(* CODESYS project Tc3_McCoordinatedMotion.library
   TcLibraryId: Beckhoff Automation GmbH|Tc3_McCoordinatedMotion|4.0.17.0
   Company: Beckhoff Automation GmbH
   Title: Tc3_McCoordinatedMotion
   Placeholder: Tc3_McCoordinatedMotion
   Version: 4.0.17.0

Project tree, tasks and I/O mapping:
  libraries: Tc2_MC2, * (Beckhoff Automation GmbH); Tc3_Mc3Definitions, 4.0.17.0 (Beckhoff Automation GmbH); Tc3_Physics, 4.0.17.0 (Beckhoff Automation GmbH)
  POUs/
    Administrative/
      function ACSIDX_TO_IDENTINGROUP [ST]
      function MCSAXISTYPE_TO_IDENTINGROUP [ST]
      function MCSIDX_TO_IDENTINGROUP [ST]
      function block MC_AddAxisToGroup [ST]: FB_init, FB_exit
      function block MC_GroupDisable [ST]: FB_init, FB_exit
      function block MC_GroupEnable [ST]: FB_init, FB_exit
      function block MC_GroupReadError [ST]: FB_init, FB_exit
      function block MC_GroupReadStatus [ST]: FB_init, FB_exit
      function block MC_GroupReadTrajectoryInformation [ST]: FB_init, FB_exit
      function block MC_GroupReset [ST]: FB_init, FB_exit
      function block MC_GroupSetOverride [ST]: FB_init, FB_exit
      function block MC_GroupSetSetpointSource [ST]: FB_init, FB_exit
      function block MC_RemoveAxisFromGroup [ST]: FB_init, FB_exit
      function block MC_SetCoordinateTransform [ST]: FB_init, FB_exit
      function block MC_SetCoordinateTransformPreparation [ST]: FB_init, FB_exit
      function block MC_TrackConveyorBelt [ST]: FB_init, FB_exit
      function block MC_UngroupAllAxes [ST]: FB_init, FB_exit
      function UDINT_TO_IDENTINGROUP [ST]
    Motion/
      function block MC_MovePath [ST]: FB_init, FB_exit
      function block MC_BlockerPreparation [ST]: FB_init, FB_exit
      function block MC_DwellTimePreparation [ST]: FB_init, FB_exit
      function block MC_GroupHalt [ST]: FB_init, FB_exit
      function block MC_GroupStop [ST]: FB_init, FB_exit
      function block MC_MoveBlendingPreparation [ST]: FB_init, FB_exit
      function block MC_MoveCircularAbsolutePreparation [ST]: FB_init, FB_exit
      function block MC_GroupReadBlockerStatus [ST]: FB_init, FB_exit
      function block MC_MoveDirectPreparation [ST]: FB_init, FB_exit
      function block MC_MoveLinearAbsolutePreparation [ST]: FB_init, FB_exit
      function block MC_ReleaseBlocker [ST]: FB_init, FB_exit
      function block MC_CalcTrafo [ST]: FB_init, FB_exit
  DUTs/
    function block MC_PATH_DATA_REF [ST]: ClearPath, FB_init, FB_exit
    data type AXES_GROUP_REF
    data type IDENT_IN_GROUP_REF
    Enums/
      data type MC_MCS_AXIS_TYPE
      data type MC_CIRC_MODE
      data type MC_CIRC_PATHCHOICE
      data type MC_TRANSITION_MODE
      data type ECmSetpointSource
      data type ETrackingSyncPosStrategy
    data type MC_COORD_REF
    data type MC_TRAJECTORY_ENTRY
    CalcTrafo/
      data type E_CalcTrafoMetaInfoScara
      data type E_CalcTrafoMetaInfo5DType1
      data type U_CalcTrafoMetaInfo
  GVLs/
    global variables GVL
  Version/
    global variables Global_Version
*)

// DUTs/AXES_GROUP_REF
(* Contains the information passed between Nc and Plc for each group. *)
{attribute 'TcIecLibraryType'}
{attribute 'Namespace' := 'Tc3_McCoordinatedMotion'}
TYPE AXES_GROUP_REF : 
	STRUCT
		(* Data from PLC to MC. *)
		{attribute 'GUID' := '0E2E3852-A98C-4AF3-81E2-209EE128940C'}
		{attribute 'Namespace' := 'MC'}
		PlcToNc AT %Q* : MC.CDT_PLCTOMC_GROUP;
		(* Data from MC to PLC. *)
		{attribute 'GUID' := '467F4325-10DF-4BC1-88DD-E8240EB4F8E3'}
		{attribute 'Namespace' := 'MC'}
		NcToPlc AT %I* : MC.CDT_MCTOPLC_GROUP;
	END_STRUCT
END_TYPE

// DUTs/IDENT_IN_GROUP_REF
{attribute 'TcIecLibraryType'}
{attribute 'Namespace' := 'Tc3_McCoordinatedMotion'}
TYPE IDENT_IN_GROUP_REF : Tc3_Physics.CoordinateType;
END_TYPE

// DUTs/MC_COORD_REF
{attribute 'TcIecLibraryType'}
{attribute 'Namespace' := 'Tc3_McCoordinatedMotion'}
TYPE MC_COORD_REF : GLOBAL.OTCID;
END_TYPE

// DUTs/MC_TRAJECTORY_ENTRY
{attribute 'TcIecLibraryType'}
{attribute 'Namespace' := 'Tc3_McCoordinatedMotion'}
TYPE MC_TRAJECTORY_ENTRY : 
	STRUCT
		InvokeId : UDINT;
		Active : BOOL;
		 {attribute 'hide'}
		_reserved1 : ARRAY [1..3] OF USINT;
		RemainingCartesianLength : LREAL;
		RemainingDuration : LREAL;
	END_STRUCT
END_TYPE

// DUTs/Enums/MC_MCS_AXIS_TYPE
{attribute 'TcIecLibraryType'}
{attribute 'Namespace' := 'Tc3_McCoordinatedMotion'}
{attribute 'hide'}
TYPE MC_MCS_AXIS_TYPE : (mcAxisTypeMcsX:=17, mcAxisTypeMcsY:=33, mcAxisTypeMcsZ:=49, mcAxisTypeMcsA1:=65, mcAxisTypeMcsA2:=66, mcAxisTypeMcsA3:=67, mcAxisTypeMcsB1:=81, mcAxisTypeMcsB2:=82, mcAxisTypeMcsB3:=83, mcAxisTypeMcsC1:=97, mcAxisTypeMcsC2:=98, mcAxisTypeMcsC3:=99) UDINT;
END_TYPE

// DUTs/Enums/MC_CIRC_MODE
{attribute 'TcIecLibraryType'}
{attribute 'Namespace' := 'Tc3_McCoordinatedMotion'}
TYPE MC_CIRC_MODE : (mcCircModeInvalid:=0, mcCircModeBorder:=8192, mcCircModeCenter:=8193, mcCircModeRadius:=8194) UINT;
END_TYPE

// DUTs/Enums/MC_CIRC_PATHCHOICE
{attribute 'TcIecLibraryType'}
{attribute 'Namespace' := 'Tc3_McCoordinatedMotion'}
TYPE MC_CIRC_PATHCHOICE : (mcCircPathChoiceClockwise:=12288, mcCircPathChoiceCounterClockwise:=12289, mcCircPathChoiceShortSegment:=12290, mcCircPathChoiceLongSegment:=12291) UINT;
END_TYPE

// DUTs/Enums/MC_TRANSITION_MODE
{attribute 'TcIecLibraryType'}
{attribute 'Namespace' := 'Tc3_McCoordinatedMotion'}
TYPE MC_TRANSITION_MODE : (mcTransModeNone:=4096, mcTransModeStartVelocity:=4097, mcTransModeConstantVelocity:=4098, mcTransModeCornerDistance:=4099, mcTransModeMaxCornerDeviation:=4100, mcTransModeCornerDistanceAdvanced:=4106) UINT;
END_TYPE

// DUTs/Enums/ECmSetpointSource
{attribute 'TcIecLibraryType'}
{attribute 'Namespace' := 'Tc3_McCoordinatedMotion'}
{attribute 'qualified_only'}
TYPE ECmSetpointSource : (Group:=1, MCS:=2, ACS:=3) UINT;
END_TYPE

// DUTs/Enums/ETrackingSyncPosStrategy
{attribute 'TcIecLibraryType'}
{attribute 'Namespace' := 'Tc3_McCoordinatedMotion'}
{attribute 'hide'}
{attribute 'qualified_only'}
TYPE ETrackingSyncPosStrategy : (FastestSync:=0, ObjectPos:=1) UINT;
END_TYPE

// DUTs/CalcTrafo/E_CalcTrafoMetaInfoScara
{attribute 'TcIecLibraryType'}
{attribute 'Namespace' := 'Tc3_McCoordinatedMotion'}
TYPE E_CalcTrafoMetaInfoScara : (scaraLeftArm:=1, scaraRightArm:=2, scaraActualConfig:=3) WORD;
END_TYPE

// DUTs/CalcTrafo/E_CalcTrafoMetaInfo5DType1
{attribute 'TcIecLibraryType'}
{attribute 'Namespace' := 'Tc3_McCoordinatedMotion'}
TYPE E_CalcTrafoMetaInfo5DType1 : (
	d5Type1Quad14:=1, 	(* M3: -90..90 and TCP in same quadrants *)
	d5Type1Quad23:=2, 	(* M3: -90..90 and TCP OUTSIDE these quadrants *)
	d5Type1ActualConfig:=3
) WORD;
END_TYPE

// DUTs/CalcTrafo/U_CalcTrafoMetaInfo
{attribute 'TcIecLibraryType'}
{attribute 'Namespace' := 'Tc3_McCoordinatedMotion'}
TYPE U_CalcTrafoMetaInfo : 
	UNION
		aData : ARRAY [1..4] OF UDINT;
		{attribute 'GUID' := '22B37A1B-3FA1-4BF4-9362-FB65E805A05C'}
		{attribute 'Namespace' := 'Tc3_McCoordinatedMotion'}
		eScara : E_CalcTrafoMetaInfoScara;
		{attribute 'GUID' := '8B943ECD-E6C5-437F-BECC-C5910C2E0300'}
		{attribute 'Namespace' := 'Tc3_McCoordinatedMotion'}
		e5dType1 : E_CalcTrafoMetaInfo5DType1;
	END_UNION
END_TYPE

// GVLs/GVL
{attribute 'external_name' := 'GVL_GUID_711467BC_BF56_4818_B36B_80DF8CEC86B5'}
{attribute 'Namespace' := 'Tc3_McCoordinatedMotion'}
VAR_GLOBAL
	MCS_X	:	IDENT_IN_GROUP_REF := MCSAXISTYPE_TO_IDENTINGROUP(mcAxisTypeMcsX);
	MCS_Y	:	IDENT_IN_GROUP_REF := MCSAXISTYPE_TO_IDENTINGROUP(mcAxisTypeMcsY);
	MCS_Z	:	IDENT_IN_GROUP_REF := MCSAXISTYPE_TO_IDENTINGROUP(mcAxisTypeMcsZ);
	MCS_A1	:	IDENT_IN_GROUP_REF := MCSAXISTYPE_TO_IDENTINGROUP(mcAxisTypeMcsA1);
	MCS_A2	:	IDENT_IN_GROUP_REF := MCSAXISTYPE_TO_IDENTINGROUP(mcAxisTypeMcsA2);
	MCS_A3	:	IDENT_IN_GROUP_REF := MCSAXISTYPE_TO_IDENTINGROUP(mcAxisTypeMcsA3);
	MCS_B1	:	IDENT_IN_GROUP_REF := MCSAXISTYPE_TO_IDENTINGROUP(mcAxisTypeMcsB1);
	MCS_B2	:	IDENT_IN_GROUP_REF := MCSAXISTYPE_TO_IDENTINGROUP(mcAxisTypeMcsB2);
	MCS_B3	:	IDENT_IN_GROUP_REF := MCSAXISTYPE_TO_IDENTINGROUP(mcAxisTypeMcsB3);
	MCS_C1	:	IDENT_IN_GROUP_REF := MCSAXISTYPE_TO_IDENTINGROUP(mcAxisTypeMcsC1);
	MCS_C2	:	IDENT_IN_GROUP_REF := MCSAXISTYPE_TO_IDENTINGROUP(mcAxisTypeMcsC2);
	MCS_C3	:	IDENT_IN_GROUP_REF := MCSAXISTYPE_TO_IDENTINGROUP(mcAxisTypeMcsC3);
	ADDAX1	:	IDENT_IN_GROUP_REF := UDINT_TO_IDENTINGROUP(1);
	ADDAX2	:	IDENT_IN_GROUP_REF := UDINT_TO_IDENTINGROUP(2);
	ADDAX3	:	IDENT_IN_GROUP_REF := UDINT_TO_IDENTINGROUP(3);
	ADDAX4	:	IDENT_IN_GROUP_REF := UDINT_TO_IDENTINGROUP(4);
	ADDAX5	:	IDENT_IN_GROUP_REF := UDINT_TO_IDENTINGROUP(5);
	ADDAX6	:	IDENT_IN_GROUP_REF := UDINT_TO_IDENTINGROUP(6);
	ADDAX7	:	IDENT_IN_GROUP_REF := UDINT_TO_IDENTINGROUP(7);
	ADDAX8	:	IDENT_IN_GROUP_REF := UDINT_TO_IDENTINGROUP(8);
	ACS1	:	IDENT_IN_GROUP_REF := ACSIDX_TO_IDENTINGROUP(1);
	ACS2	:	IDENT_IN_GROUP_REF := ACSIDX_TO_IDENTINGROUP(2);
	ACS3	:	IDENT_IN_GROUP_REF := ACSIDX_TO_IDENTINGROUP(3);
	ACS4	:	IDENT_IN_GROUP_REF := ACSIDX_TO_IDENTINGROUP(4);
	ACS5	:	IDENT_IN_GROUP_REF := ACSIDX_TO_IDENTINGROUP(5);
	ACS6	:	IDENT_IN_GROUP_REF := ACSIDX_TO_IDENTINGROUP(6);
END_VAR

// Version/Global_Version
{attribute 'TcGenerated'}
// This function has been automatically generated from the project information.
VAR_GLOBAL CONSTANT
	{attribute 'const_non_replaced'}
	{attribute 'linkalways'}
	stLibVersion_Tc3_McCoordinatedMotion : ST_LibVersion := (iMajor := 4, iMinor := 0, iBuild := 17, iRevision := 0, nFlags := 0, sVersion := '4.0.17.0');
	{attribute 'const_non_replaced'}
	{attribute 'linkalways'}
	sLibraryId_Tc3_McCoordinatedMotion : String := 'Beckhoff Automation GmbH|Tc3_McCoordinatedMotion|4.0.17.0';
END_VAR

// DUTs/MC_PATH_DATA_REF

{attribute 'c++_compatible'}
{attribute 'external_name' := 'MC_PATH_DATA_REF_GUID_C9AD990F_1976_3217_E176_0481FCAF8F1C'}
{attribute 'TcIecLibraryType'}
{attribute 'hide_all_locals'}
FUNCTION_BLOCK MC_PATH_DATA_REF
VAR_OUTPUT
	FilledRows : UDINT;
	OccupiedBuffer : UDINT;
END_VAR
VAR
	{attribute 'GUID' := '18071995-0000-0000-0000-000000000018'}
	StreamHdr : GLOBAL.PVOID;
	BufferSize : UDINT;
	 {attribute 'hide'}
	_reserved1 : UINT_0_32;
	{attribute 'GUID' := '18071995-0000-0000-0000-000000000018'}
	Top : GLOBAL.PVOID;
	{attribute 'GUID' := '18071995-0000-0000-0000-000000000019'}
	InternalError : GLOBAL.HRESULT;
END_VAR

{attribute 'TcTypeSystem'}

METHOD ClearPath
END_METHOD

{attribute 'TcTypeSystem'}

(* Internal method *)
{attribute 'hide'}
METHOD FB_init : BOOL
VAR_INPUT
	(*  if TRUE, the retain variables are initialized (warm start / cold start) *)
	bInitRetains : BOOL;
	(*  if TRUE, the instance afterwards gets moved into the copy code (online change) *)
	bInCopyCode : BOOL;
	(*  buffer to store elements of path, use ADR(...) *)
	{attribute 'GUID' := '18071995-0000-0000-0000-000000000018'}
	pBuffer : GLOBAL.PVOID;
	(*  size of buffer (in Bytes), use SIZEOF(...) *)
	nBufferSize : UDINT;
END_VAR
END_METHOD

{attribute 'TcTypeSystem'}

(* Internal method *)
{attribute 'hide'}
METHOD FB_exit : BOOL
VAR_INPUT
	(*  if TRUE, the exit method is called for exiting an instance that is copied afterwards (online change). *)
	bInCopyCode : BOOL;
END_VAR
END_METHOD

END_FUNCTION_BLOCK

// POUs/Administrative/ACSIDX_TO_IDENTINGROUP
{attribute 'TcIecLibraryType'}
{attribute 'external_name' := 'ACSIDX_TO_IDENTINGROUP_GUID_B36A848B_1747_3CA7_C03B_4EEFE5351486'}
{attribute 'Namespace' := 'Tc3_McCoordinatedMotion'}
{attribute 'hide'}
FUNCTION ACSIDX_TO_IDENTINGROUP : IDENT_IN_GROUP_REF
VAR_INPUT
	AcsIndex	:	UDINT;	(* Index in Axis Coordinate System (relevant for Kinematics) *)
END_VAR

END_FUNCTION

// POUs/Administrative/MCSAXISTYPE_TO_IDENTINGROUP
{attribute 'TcIecLibraryType'}
{attribute 'external_name' := 'MCSAXISTYPE_TO_IDENTINGROUP_GUID_6F5B7E7F_56A6_3E32_D091_CE95291E5C23'}
{attribute 'Namespace' := 'Tc3_McCoordinatedMotion'}
{attribute 'hide'}
FUNCTION MCSAXISTYPE_TO_IDENTINGROUP : IDENT_IN_GROUP_REF
VAR_INPUT
	AxisType	:	MC_MCS_AXIS_TYPE;	(* Axis Interpretation in Machine Coordinate System *)
END_VAR

END_FUNCTION

// POUs/Administrative/MCSIDX_TO_IDENTINGROUP
{attribute 'TcIecLibraryType'}
{attribute 'external_name' := 'MCSIDX_TO_IDENTINGROUP_GUID_41217B1F_38B5_340B_DB7E_B8FA4F687802'}
{attribute 'Namespace' := 'Tc3_McCoordinatedMotion'}
{attribute 'hide'}
FUNCTION MCSIDX_TO_IDENTINGROUP : IDENT_IN_GROUP_REF
VAR_INPUT
	McsIndex	:	UDINT;	(* Index in Machine Coordinate System *)
END_VAR

END_FUNCTION

// POUs/Administrative/MC_AddAxisToGroup

{attribute 'c++_compatible'}
{attribute 'external_name' := 'MC_AddAxisToGroup_GUID_60E0109C_AD81_3D18_D844_0BD44DAFCDF2'}
{attribute 'TcIecLibraryType'}
{attribute 'hide_all_locals'}
FUNCTION_BLOCK MC_AddAxisToGroup
VAR_IN_OUT
	(* B *)
	{attribute 'GUID' := 'EE658783-7533-4695-9194-9C08CBE11A9C'}
	{attribute 'Namespace' := 'Tc3_McCoordinatedMotion'}
	AxesGroup : AXES_GROUP_REF;
	(* B *)
	{attribute 'GUID' := '796382E2-8BB1-4613-AF21-647CD1FFE3C7'}
	{attribute 'Namespace' := 'Tc2_MC2'}
	Axis : Tc2_MC2.AXIS_REF;
END_VAR
VAR_INPUT
	(* B *)
	Execute : BOOL;
END_VAR
VAR
	 {attribute 'hide'}
	_reserved1 : UINT_24_56;
END_VAR
VAR_INPUT
	(* E *)
	{attribute 'GUID' := 'CB1E2F74-F48F-4B08-86F0-C3153004E775'}
	{attribute 'Namespace' := 'Tc3_McCoordinatedMotion'}
	IdentInGroup : IDENT_IN_GROUP_REF;
END_VAR
VAR_OUTPUT
	(* B *)
	Done : BOOL;
	(* E *)
	Busy : BOOL;
	(* B *)
	Error : BOOL;
END_VAR
VAR
	 {attribute 'hide'}
	_reserved2 : USINT;
END_VAR
VAR_OUTPUT
	(* E *)
	ErrorId : UDINT;
END_VAR
VAR
	InternalFBState : ARRAY [1..16] OF ULINT;
END_VAR

{attribute 'TcTypeSystem'}

(* Internal method *)
{attribute 'hide'}
METHOD FB_init : BOOL
VAR_INPUT
	(*  if TRUE, the retain variables are initialized (warm start / cold start) *)
	bInitRetains : BOOL;
	(*  if TRUE, the instance afterwards gets moved into the copy code (online change) *)
	bInCopyCode : BOOL;
END_VAR
END_METHOD

{attribute 'TcTypeSystem'}

(* Internal method *)
{attribute 'hide'}
METHOD FB_exit : BOOL
VAR_INPUT
	(*  if TRUE, the exit method is called for exiting an instance that is copied afterwards (online change). *)
	bInCopyCode : BOOL;
END_VAR
END_METHOD

END_FUNCTION_BLOCK

// POUs/Administrative/MC_GroupDisable

{attribute 'c++_compatible'}
{attribute 'external_name' := 'MC_GroupDisable_GUID_87A0F0BD_AB84_365F_DF81_18084A213C76'}
{attribute 'TcIecLibraryType'}
{attribute 'hide_all_locals'}
FUNCTION_BLOCK MC_GroupDisable
VAR_IN_OUT
	(* B *)
	{attribute 'GUID' := 'EE658783-7533-4695-9194-9C08CBE11A9C'}
	{attribute 'Namespace' := 'Tc3_McCoordinatedMotion'}
	AxesGroup : AXES_GROUP_REF;
END_VAR
VAR_INPUT
	(* B *)
	Execute : BOOL;
END_VAR
VAR_OUTPUT
	(* B *)
	Done : BOOL;
	(* E *)
	Busy : BOOL;
	(* B *)
	Error : BOOL;
	(* E *)
	ErrorId : UDINT;
END_VAR
VAR
	InternalFBState : ARRAY [1..16] OF ULINT;
END_VAR

{attribute 'TcTypeSystem'}

(* Internal method *)
{attribute 'hide'}
METHOD FB_init : BOOL
VAR_INPUT
	(*  if TRUE, the retain variables are initialized (warm start / cold start) *)
	bInitRetains : BOOL;
	(*  if TRUE, the instance afterwards gets moved into the copy code (online change) *)
	bInCopyCode : BOOL;
END_VAR
END_METHOD

{attribute 'TcTypeSystem'}

(* Internal method *)
{attribute 'hide'}
METHOD FB_exit : BOOL
VAR_INPUT
	(*  if TRUE, the exit method is called for exiting an instance that is copied afterwards (online change). *)
	bInCopyCode : BOOL;
END_VAR
END_METHOD

END_FUNCTION_BLOCK

// POUs/Administrative/MC_GroupEnable

{attribute 'c++_compatible'}
{attribute 'external_name' := 'MC_GroupEnable_GUID_7A2FA050_093A_3C93_F1B8_5490C7CC913F'}
{attribute 'TcIecLibraryType'}
{attribute 'hide_all_locals'}
FUNCTION_BLOCK MC_GroupEnable
VAR_IN_OUT
	(* B *)
	{attribute 'GUID' := 'EE658783-7533-4695-9194-9C08CBE11A9C'}
	{attribute 'Namespace' := 'Tc3_McCoordinatedMotion'}
	AxesGroup : AXES_GROUP_REF;
END_VAR
VAR_INPUT
	(* B *)
	Execute : BOOL;
END_VAR
VAR_OUTPUT
	(* B *)
	Done : BOOL;
	(* E *)
	Busy : BOOL;
	(* B *)
	Error : BOOL;
	(* E *)
	ErrorId : UDINT;
END_VAR
VAR
	InternalFBState : ARRAY [1..16] OF ULINT;
END_VAR

{attribute 'TcTypeSystem'}

(* Internal method *)
{attribute 'hide'}
METHOD FB_init : BOOL
VAR_INPUT
	(*  if TRUE, the retain variables are initialized (warm start / cold start) *)
	bInitRetains : BOOL;
	(*  if TRUE, the instance afterwards gets moved into the copy code (online change) *)
	bInCopyCode : BOOL;
END_VAR
END_METHOD

{attribute 'TcTypeSystem'}

(* Internal method *)
{attribute 'hide'}
METHOD FB_exit : BOOL
VAR_INPUT
	(*  if TRUE, the exit method is called for exiting an instance that is copied afterwards (online change). *)
	bInCopyCode : BOOL;
END_VAR
END_METHOD

END_FUNCTION_BLOCK

// POUs/Administrative/MC_GroupReadError

{attribute 'c++_compatible'}
{attribute 'external_name' := 'MC_GroupReadError_GUID_B8E629EB_C7F2_3B02_D695_647A427CC122'}
{attribute 'TcIecLibraryType'}
{attribute 'hide_all_locals'}
FUNCTION_BLOCK MC_GroupReadError
VAR_IN_OUT
	(* B *)
	{attribute 'GUID' := 'EE658783-7533-4695-9194-9C08CBE11A9C'}
	{attribute 'Namespace' := 'Tc3_McCoordinatedMotion'}
	AxesGroup : AXES_GROUP_REF;
END_VAR
VAR_INPUT
	(* B *)
	Enable : BOOL;
END_VAR
VAR_OUTPUT
	(* B *)
	Valid : BOOL;
	(* E *)
	Busy : BOOL;
	(* B *)
	Error : BOOL;
	(* E *)
	ErrorId : UDINT;
	(* E *)
	GroupErrorId : UDINT;
END_VAR
VAR
END_VAR

{attribute 'TcTypeSystem'}

(* Internal method *)
{attribute 'hide'}
METHOD FB_init : BOOL
VAR_INPUT
	(*  if TRUE, the retain variables are initialized (warm start / cold start) *)
	bInitRetains : BOOL;
	(*  if TRUE, the instance afterwards gets moved into the copy code (online change) *)
	bInCopyCode : BOOL;
END_VAR
END_METHOD

{attribute 'TcTypeSystem'}

(* Internal method *)
{attribute 'hide'}
METHOD FB_exit : BOOL
VAR_INPUT
	(*  if TRUE, the exit method is called for exiting an instance that is copied afterwards (online change). *)
	bInCopyCode : BOOL;
END_VAR
END_METHOD

END_FUNCTION_BLOCK

// POUs/Administrative/MC_GroupReadStatus

{attribute 'c++_compatible'}
{attribute 'external_name' := 'MC_GroupReadStatus_GUID_BD62E39C_B8A7_357C_C275_26E3AC2C5659'}
{attribute 'TcIecLibraryType'}
{attribute 'hide_all_locals'}
FUNCTION_BLOCK MC_GroupReadStatus
VAR_IN_OUT
	(* B *)
	{attribute 'GUID' := 'EE658783-7533-4695-9194-9C08CBE11A9C'}
	{attribute 'Namespace' := 'Tc3_McCoordinatedMotion'}
	AxesGroup : AXES_GROUP_REF;
END_VAR
VAR_INPUT
	(* B *)
	Enable : BOOL;
END_VAR
VAR_OUTPUT
	(* B *)
	Valid : BOOL;
	(* E *)
	Busy : BOOL;
	(* E *)
	GroupMoving : BOOL;
	(* E *)
	GroupHoming : BOOL;
	(* E *)
	GroupErrorStop : BOOL;
	(* E *)
	GroupNotReady : BOOL;
	(* E *)
	GroupStandby : BOOL;
	(* E *)
	GroupStopping : BOOL;
	(* E *)
	GroupDisabled : BOOL;
	(* E *)
	AllAxesStanding : BOOL;
	(* E *)
	{attribute 'hide'}
	ConstantVelocity : BOOL;
	(* E *)
	{attribute 'hide'}
	Accelerating : BOOL;
	(* E *)
	{attribute 'hide'}
	Decelerating : BOOL;
	(* E *)
	InPosition : BOOL;
	(* B *)
	Error : BOOL;
	(* E *)
	ErrorId : UDINT;
END_VAR
VAR
END_VAR

{attribute 'TcTypeSystem'}

(* Internal method *)
{attribute 'hide'}
METHOD FB_init : BOOL
VAR_INPUT
	(*  if TRUE, the retain variables are initialized (warm start / cold start) *)
	bInitRetains : BOOL;
	(*  if TRUE, the instance afterwards gets moved into the copy code (online change) *)
	bInCopyCode : BOOL;
END_VAR
END_METHOD

{attribute 'TcTypeSystem'}

(* Internal method *)
{attribute 'hide'}
METHOD FB_exit : BOOL
VAR_INPUT
	(*  if TRUE, the exit method is called for exiting an instance that is copied afterwards (online change). *)
	bInCopyCode : BOOL;
END_VAR
END_METHOD

END_FUNCTION_BLOCK

// POUs/Administrative/MC_GroupReadTrajectoryInformation

{attribute 'c++_compatible'}
{attribute 'external_name' := 'MC_GroupReadTrajectoryInformation_GUID_31A53C6A_DFF7_3689_C5EB_3A3FD6ED5762'}
{attribute 'TcIecLibraryType'}
{attribute 'hide_all_locals'}
FUNCTION_BLOCK MC_GroupReadTrajectoryInformation
VAR_IN_OUT
	(* B *)
	{attribute 'GUID' := 'EE658783-7533-4695-9194-9C08CBE11A9C'}
	{attribute 'Namespace' := 'Tc3_McCoordinatedMotion'}
	AxesGroup : AXES_GROUP_REF;
END_VAR
VAR_INPUT
	(* B *)
	Enable : BOOL;
END_VAR
VAR_OUTPUT
	(* B *)
	Valid : BOOL;
	(* B *)
	Error : BOOL;
END_VAR
VAR
	 {attribute 'hide'}
	_reserved1 : USINT;
END_VAR
VAR_OUTPUT
	(* E *)
	ErrorId : UDINT;
	(* E *)
	EntryCount : UDINT;
END_VAR
VAR
	 {attribute 'hide'}
	_reserved2 : UDINT;
END_VAR
VAR_OUTPUT
	(* E *)
	{attribute 'GUID' := 'F7E5A6B8-C9D0-4E1F-AA3B-4C5D6E7F8091'}
	{attribute 'Namespace' := 'Tc3_McCoordinatedMotion'}
	Entries : ARRAY [1..10] OF MC_TRAJECTORY_ENTRY;
END_VAR
VAR
END_VAR

{attribute 'TcTypeSystem'}

(* Internal method *)
{attribute 'hide'}
METHOD FB_init : BOOL
VAR_INPUT
	(*  if TRUE, the retain variables are initialized (warm start / cold start) *)
	bInitRetains : BOOL;
	(*  if TRUE, the instance afterwards gets moved into the copy code (online change) *)
	bInCopyCode : BOOL;
END_VAR
END_METHOD

{attribute 'TcTypeSystem'}

(* Internal method *)
{attribute 'hide'}
METHOD FB_exit : BOOL
VAR_INPUT
	(*  if TRUE, the exit method is called for exiting an instance that is copied afterwards (online change). *)
	bInCopyCode : BOOL;
END_VAR
END_METHOD

END_FUNCTION_BLOCK

// POUs/Administrative/MC_GroupReset

{attribute 'c++_compatible'}
{attribute 'external_name' := 'MC_GroupReset_GUID_3781F46E_6B77_3CFC_E33A_C347CF00C0C8'}
{attribute 'TcIecLibraryType'}
{attribute 'hide_all_locals'}
FUNCTION_BLOCK MC_GroupReset
VAR_IN_OUT
	(* B *)
	{attribute 'GUID' := 'EE658783-7533-4695-9194-9C08CBE11A9C'}
	{attribute 'Namespace' := 'Tc3_McCoordinatedMotion'}
	AxesGroup : AXES_GROUP_REF;
END_VAR
VAR_INPUT
	(* B *)
	Execute : BOOL;
END_VAR
VAR_OUTPUT
	(* B *)
	Done : BOOL;
	(* E *)
	Busy : BOOL;
	(* B *)
	Error : BOOL;
	(* E *)
	ErrorId : UDINT;
END_VAR
VAR
	InternalFBState : ARRAY [1..16] OF ULINT;
END_VAR

{attribute 'TcTypeSystem'}

(* Internal method *)
{attribute 'hide'}
METHOD FB_init : BOOL
VAR_INPUT
	(*  if TRUE, the retain variables are initialized (warm start / cold start) *)
	bInitRetains : BOOL;
	(*  if TRUE, the instance afterwards gets moved into the copy code (online change) *)
	bInCopyCode : BOOL;
END_VAR
END_METHOD

{attribute 'TcTypeSystem'}

(* Internal method *)
{attribute 'hide'}
METHOD FB_exit : BOOL
VAR_INPUT
	(*  if TRUE, the exit method is called for exiting an instance that is copied afterwards (online change). *)
	bInCopyCode : BOOL;
END_VAR
END_METHOD

END_FUNCTION_BLOCK

// POUs/Administrative/MC_GroupSetOverride

{attribute 'c++_compatible'}
{attribute 'external_name' := 'MC_GroupSetOverride_GUID_CA3640F9_4BC4_37DE_EFFB_93C36A60C3E3'}
{attribute 'TcIecLibraryType'}
{attribute 'hide_all_locals'}
FUNCTION_BLOCK MC_GroupSetOverride
VAR_IN_OUT
	(* B *)
	{attribute 'GUID' := 'EE658783-7533-4695-9194-9C08CBE11A9C'}
	{attribute 'Namespace' := 'Tc3_McCoordinatedMotion'}
	AxesGroup : AXES_GROUP_REF;
END_VAR
VAR_INPUT
	(* B *)
	Enable : BOOL;
END_VAR
VAR
	 {attribute 'hide'}
	_reserved1 : ARRAY [1..7] OF USINT;
END_VAR
VAR_INPUT
	(* E *)
	{attribute 'GUID' := '0100FF8A-3F83-4535-990A-614CFBA4DA63'}
	{attribute 'Namespace' := 'MC'}
	VelFactor : MC.MC_LREAL;
END_VAR
VAR_OUTPUT
	(* E *)
	Enabled : BOOL;
	(* E *)
	Busy : BOOL;
	(* B *)
	Error : BOOL;
END_VAR
VAR
	 {attribute 'hide'}
	_reserved2 : USINT;
END_VAR
VAR_OUTPUT
	(* E *)
	ErrorId : UDINT;
	(* E *)
	ActualVelFactor : LREAL;
END_VAR
VAR
END_VAR

{attribute 'TcTypeSystem'}

(* Internal method *)
{attribute 'hide'}
METHOD FB_init : BOOL
VAR_INPUT
	(*  if TRUE, the retain variables are initialized (warm start / cold start) *)
	bInitRetains : BOOL;
	(*  if TRUE, the instance afterwards gets moved into the copy code (online change) *)
	bInCopyCode : BOOL;
END_VAR
END_METHOD

{attribute 'TcTypeSystem'}

(* Internal method *)
{attribute 'hide'}
METHOD FB_exit : BOOL
VAR_INPUT
	(*  if TRUE, the exit method is called for exiting an instance that is copied afterwards (online change). *)
	bInCopyCode : BOOL;
END_VAR
END_METHOD

END_FUNCTION_BLOCK

// POUs/Administrative/MC_GroupSetSetpointSource

{attribute 'c++_compatible'}
{attribute 'external_name' := 'MC_GroupSetSetpointSource_GUID_5F373C6C_C746_32C0_F0B7_E48FC09F6070'}
{attribute 'TcIecLibraryType'}
{attribute 'hide_all_locals'}
FUNCTION_BLOCK MC_GroupSetSetpointSource
VAR_IN_OUT
	(* B *)
	{attribute 'GUID' := 'EE658783-7533-4695-9194-9C08CBE11A9C'}
	{attribute 'Namespace' := 'Tc3_McCoordinatedMotion'}
	AxesGroup : AXES_GROUP_REF;
END_VAR
VAR_INPUT
	(* B *)
	Execute : BOOL;
END_VAR
VAR
	 {attribute 'hide'}
	_reserved1 : USINT;
END_VAR
VAR_INPUT
	(* E *)
	{attribute 'GUID' := 'D0A61B70-69A5-45AB-898B-011D56402A97'}
	{attribute 'Namespace' := 'Tc3_McCoordinatedMotion'}
	SetpointSource : ECmSetpointSource;
END_VAR
VAR_OUTPUT
	(* B *)
	Done : BOOL;
	(* E *)
	Busy : BOOL;
	(* B *)
	Error : BOOL;
END_VAR
VAR
	 {attribute 'hide'}
	_reserved2 : USINT;
END_VAR
VAR_OUTPUT
	(* E *)
	ErrorId : UDINT;
END_VAR
VAR
	 {attribute 'hide'}
	_reserved3 : UDINT;
	InternalFBState : ARRAY [1..16] OF ULINT;
END_VAR

{attribute 'TcTypeSystem'}

(* Internal method *)
{attribute 'hide'}
METHOD FB_init : BOOL
VAR_INPUT
	(*  if TRUE, the retain variables are initialized (warm start / cold start) *)
	bInitRetains : BOOL;
	(*  if TRUE, the instance afterwards gets moved into the copy code (online change) *)
	bInCopyCode : BOOL;
END_VAR
END_METHOD

{attribute 'TcTypeSystem'}

(* Internal method *)
{attribute 'hide'}
METHOD FB_exit : BOOL
VAR_INPUT
	(*  if TRUE, the exit method is called for exiting an instance that is copied afterwards (online change). *)
	bInCopyCode : BOOL;
END_VAR
END_METHOD

END_FUNCTION_BLOCK

// POUs/Administrative/MC_RemoveAxisFromGroup

{attribute 'c++_compatible'}
{attribute 'external_name' := 'MC_RemoveAxisFromGroup_GUID_22EDF44C_D9C3_3A6F_FBE1_FFD3C2A62A3E'}
{attribute 'TcIecLibraryType'}
{attribute 'hide_all_locals'}
FUNCTION_BLOCK MC_RemoveAxisFromGroup
VAR_IN_OUT
	(* B *)
	{attribute 'GUID' := 'EE658783-7533-4695-9194-9C08CBE11A9C'}
	{attribute 'Namespace' := 'Tc3_McCoordinatedMotion'}
	AxesGroup : AXES_GROUP_REF;
END_VAR
VAR_INPUT
	(* B *)
	Execute : BOOL;
END_VAR
VAR
	 {attribute 'hide'}
	_reserved1 : ARRAY [1..7] OF USINT;
END_VAR
VAR_INPUT
	(* B *)
	{attribute 'GUID' := 'CB1E2F74-F48F-4B08-86F0-C3153004E775'}
	{attribute 'Namespace' := 'Tc3_McCoordinatedMotion'}
	IdentInGroup : IDENT_IN_GROUP_REF;
END_VAR
VAR_OUTPUT
	(* B *)
	Done : BOOL;
	(* E *)
	Busy : BOOL;
	(* B *)
	Error : BOOL;
END_VAR
VAR
	 {attribute 'hide'}
	_reserved2 : USINT;
END_VAR
VAR_OUTPUT
	(* E *)
	ErrorId : UDINT;
END_VAR
VAR
	InternalFBState : ARRAY [1..16] OF ULINT;
END_VAR

{attribute 'TcTypeSystem'}

(* Internal method *)
{attribute 'hide'}
METHOD FB_init : BOOL
VAR_INPUT
	(*  if TRUE, the retain variables are initialized (warm start / cold start) *)
	bInitRetains : BOOL;
	(*  if TRUE, the instance afterwards gets moved into the copy code (online change) *)
	bInCopyCode : BOOL;
END_VAR
END_METHOD

{attribute 'TcTypeSystem'}

(* Internal method *)
{attribute 'hide'}
METHOD FB_exit : BOOL
VAR_INPUT
	(*  if TRUE, the exit method is called for exiting an instance that is copied afterwards (online change). *)
	bInCopyCode : BOOL;
END_VAR
END_METHOD

END_FUNCTION_BLOCK

// POUs/Administrative/MC_SetCoordinateTransform

{attribute 'c++_compatible'}
{attribute 'external_name' := 'MC_SetCoordinateTransform_GUID_F89D3506_B8FA_328A_EE82_986052F4EB84'}
{attribute 'TcIecLibraryType'}
{attribute 'hide_all_locals'}
FUNCTION_BLOCK MC_SetCoordinateTransform
VAR_IN_OUT
	(* B *)
	{attribute 'GUID' := 'EE658783-7533-4695-9194-9C08CBE11A9C'}
	{attribute 'Namespace' := 'Tc3_McCoordinatedMotion'}
	AxesGroup : AXES_GROUP_REF;
END_VAR
VAR_INPUT
	(* B *)
	Execute : BOOL;
END_VAR
VAR
	 {attribute 'hide'}
	_reserved1 : ARRAY [1..3] OF USINT;
END_VAR
VAR_INPUT
	(* E *)
	{attribute 'GUID' := 'E6D4F5A7-B8C9-4D0E-9F2A-3B4C5D6E7F80'}
	{attribute 'Namespace' := 'Tc3_McCoordinatedMotion'}
	CoordTransform : MC_COORD_REF;
END_VAR
VAR_OUTPUT
	(* B *)
	Done : BOOL;
	(* E *)
	Busy : BOOL;
	(* E *)
	Active : BOOL;
	(* E *)
	CommandAborted : BOOL;
	(* B *)
	Error : BOOL;
END_VAR
VAR
	 {attribute 'hide'}
	_reserved2 : ARRAY [1..3] OF USINT;
END_VAR
VAR_OUTPUT
	(* E *)
	ErrorId : UDINT;
END_VAR
VAR
	 {attribute 'hide'}
	_reserved3 : UDINT;
	InternalFBState : ARRAY [1..16] OF ULINT;
END_VAR

{attribute 'TcTypeSystem'}

(* Internal method *)
{attribute 'hide'}
METHOD FB_init : BOOL
VAR_INPUT
	(*  if TRUE, the retain variables are initialized (warm start / cold start) *)
	bInitRetains : BOOL;
	(*  if TRUE, the instance afterwards gets moved into the copy code (online change) *)
	bInCopyCode : BOOL;
END_VAR
END_METHOD

{attribute 'TcTypeSystem'}

(* Internal method *)
{attribute 'hide'}
METHOD FB_exit : BOOL
VAR_INPUT
	(*  if TRUE, the exit method is called for exiting an instance that is copied afterwards (online change). *)
	bInCopyCode : BOOL;
END_VAR
END_METHOD

END_FUNCTION_BLOCK

// POUs/Administrative/MC_SetCoordinateTransformPreparation

{attribute 'c++_compatible'}
{attribute 'external_name' := 'MC_SetCoordinateTransformPreparation_GUID_7B402EE7_D28D_32DB_F07F_69DEF823D0E8'}
{attribute 'TcIecLibraryType'}
{attribute 'hide_all_locals'}
FUNCTION_BLOCK MC_SetCoordinateTransformPreparation
VAR_IN_OUT
	(* B *)
	{attribute 'GUID' := 'C9AD990F-1976-3217-E176-0481FCAF8F1C'}
	{attribute 'Namespace' := 'Tc3_McCoordinatedMotion'}
	PathData : MC_PATH_DATA_REF;
END_VAR
VAR_INPUT
	(* E *)
	{attribute 'GUID' := 'E6D4F5A7-B8C9-4D0E-9F2A-3B4C5D6E7F80'}
	{attribute 'Namespace' := 'Tc3_McCoordinatedMotion'}
	CoordTransform : MC_COORD_REF;
END_VAR
VAR_OUTPUT
	(* B *)
	Error : BOOL;
END_VAR
VAR
	 {attribute 'hide'}
	_reserved1 : ARRAY [1..3] OF USINT;
END_VAR
VAR_OUTPUT
	(* E *)
	ErrorId : UDINT;
END_VAR
VAR
END_VAR

{attribute 'TcTypeSystem'}

(* Internal method *)
{attribute 'hide'}
METHOD FB_init : BOOL
VAR_INPUT
	(*  if TRUE, the retain variables are initialized (warm start / cold start) *)
	bInitRetains : BOOL;
	(*  if TRUE, the instance afterwards gets moved into the copy code (online change) *)
	bInCopyCode : BOOL;
END_VAR
END_METHOD

{attribute 'TcTypeSystem'}

(* Internal method *)
{attribute 'hide'}
METHOD FB_exit : BOOL
VAR_INPUT
	(*  if TRUE, the exit method is called for exiting an instance that is copied afterwards (online change). *)
	bInCopyCode : BOOL;
END_VAR
END_METHOD

END_FUNCTION_BLOCK

// POUs/Administrative/MC_TrackConveyorBelt

{attribute 'c++_compatible'}
{attribute 'external_name' := 'MC_TrackConveyorBelt_GUID_7C82869C_7BCF_3EC6_DCAE_54348C2A2EA9'}
{attribute 'TcIecLibraryType'}
{attribute 'hide_all_locals'}
FUNCTION_BLOCK MC_TrackConveyorBelt
VAR_IN_OUT
	(* B *)
	{attribute 'GUID' := 'EE658783-7533-4695-9194-9C08CBE11A9C'}
	{attribute 'Namespace' := 'Tc3_McCoordinatedMotion'}
	AxesGroup : AXES_GROUP_REF;
	(* B *)
	{attribute 'GUID' := '796382E2-8BB1-4613-AF21-647CD1FFE3C7'}
	{attribute 'Namespace' := 'Tc2_MC2'}
	ConveyorBelt : Tc2_MC2.AXIS_REF;
END_VAR
VAR_INPUT
	(* B *)
	Execute : BOOL;
END_VAR
VAR
	 {attribute 'hide'}
	_reserved1 : ARRAY [1..3] OF USINT;
END_VAR
VAR_INPUT
	(* E *)
	{attribute 'GUID' := 'E6D4F5A7-B8C9-4D0E-9F2A-3B4C5D6E7F80'}
	{attribute 'Namespace' := 'Tc3_McCoordinatedMotion'}
	CoordTransform : MC_COORD_REF;
	(* E *)
	{attribute 'GUID' := '18071995-0000-0000-0000-000000000018'}
	InitialObjectPos : GLOBAL.PVOID;
	(* E *)
	InitialObjectPosCount : UDINT;
END_VAR
VAR
	 {attribute 'hide'}
	_reserved2 : UDINT;
END_VAR
VAR_INPUT
	(* E *)
	{attribute 'GUID' := '0100FF8A-3F83-4535-990A-614CFBA4DA63'}
	{attribute 'Namespace' := 'MC'}
	MasterRefPos : MC.MC_LREAL;
	(* E *)
	{attribute 'GUID' := '0100FF8A-3F83-4535-990A-614CFBA4DA63'}
	{attribute 'Namespace' := 'MC'}
	Velocity : MC.MC_LREAL;
	(* E *)
	{attribute 'GUID' := '0100FF8A-3F83-4535-990A-614CFBA4DA63'}
	{attribute 'Namespace' := 'MC'}
	Acceleration : MC.MC_LREAL;
	(* E *)
	{attribute 'GUID' := '0100FF8A-3F83-4535-990A-614CFBA4DA63'}
	{attribute 'Namespace' := 'MC'}
	Deceleration : MC.MC_LREAL;
	(* E *)
	{attribute 'GUID' := '0100FF8A-3F83-4535-990A-614CFBA4DA63'}
	{attribute 'Namespace' := 'MC'}
	Jerk : MC.MC_LREAL;
	(* E *)
	{attribute 'hide'}
	{attribute 'GUID' := '820815FE-AACA-4B9D-9960-80212016890E'}
	{attribute 'Namespace' := 'Tc3_McCoordinatedMotion'}
	SyncPosStrategy : ETrackingSyncPosStrategy;
END_VAR
VAR_OUTPUT
	(* B *)
	InSync : BOOL;
	(* E *)
	Busy : BOOL;
	(* E *)
	Active : BOOL;
	(* E *)
	CommandAborted : BOOL;
	(* B *)
	Error : BOOL;
END_VAR
VAR
	 {attribute 'hide'}
	_reserved3 : USINT;
END_VAR
VAR_OUTPUT
	(* E *)
	ErrorId : UDINT;
END_VAR
VAR
	 {attribute 'hide'}
	_reserved4 : UDINT;
	InternalFBState : ARRAY [1..16] OF ULINT;
END_VAR

{attribute 'TcTypeSystem'}

(* Internal method *)
{attribute 'hide'}
METHOD FB_init : BOOL
VAR_INPUT
	(*  if TRUE, the retain variables are initialized (warm start / cold start) *)
	bInitRetains : BOOL;
	(*  if TRUE, the instance afterwards gets moved into the copy code (online change) *)
	bInCopyCode : BOOL;
END_VAR
END_METHOD

{attribute 'TcTypeSystem'}

(* Internal method *)
{attribute 'hide'}
METHOD FB_exit : BOOL
VAR_INPUT
	(*  if TRUE, the exit method is called for exiting an instance that is copied afterwards (online change). *)
	bInCopyCode : BOOL;
END_VAR
END_METHOD

END_FUNCTION_BLOCK

// POUs/Administrative/MC_UngroupAllAxes

{attribute 'c++_compatible'}
{attribute 'external_name' := 'MC_UngroupAllAxes_GUID_B65DD720_40E1_3BF7_DB6B_655F99D62929'}
{attribute 'TcIecLibraryType'}
{attribute 'hide_all_locals'}
FUNCTION_BLOCK MC_UngroupAllAxes
VAR_IN_OUT
	(* B *)
	{attribute 'GUID' := 'EE658783-7533-4695-9194-9C08CBE11A9C'}
	{attribute 'Namespace' := 'Tc3_McCoordinatedMotion'}
	AxesGroup : AXES_GROUP_REF;
END_VAR
VAR_INPUT
	(* B *)
	Execute : BOOL;
END_VAR
VAR_OUTPUT
	(* B *)
	Done : BOOL;
	(* E *)
	Busy : BOOL;
	(* B *)
	Error : BOOL;
	(* E *)
	ErrorId : UDINT;
END_VAR
VAR
	InternalFBState : ARRAY [1..16] OF ULINT;
END_VAR

{attribute 'TcTypeSystem'}

(* Internal method *)
{attribute 'hide'}
METHOD FB_init : BOOL
VAR_INPUT
	(*  if TRUE, the retain variables are initialized (warm start / cold start) *)
	bInitRetains : BOOL;
	(*  if TRUE, the instance afterwards gets moved into the copy code (online change) *)
	bInCopyCode : BOOL;
END_VAR
END_METHOD

{attribute 'TcTypeSystem'}

(* Internal method *)
{attribute 'hide'}
METHOD FB_exit : BOOL
VAR_INPUT
	(*  if TRUE, the exit method is called for exiting an instance that is copied afterwards (online change). *)
	bInCopyCode : BOOL;
END_VAR
END_METHOD

END_FUNCTION_BLOCK

// POUs/Administrative/UDINT_TO_IDENTINGROUP
{attribute 'TcIecLibraryType'}
{attribute 'external_name' := 'UDINT_TO_IDENTINGROUP_GUID_A56181A6_7862_387F_CCDD_ACC9D7B7D54D'}
{attribute 'Namespace' := 'Tc3_McCoordinatedMotion'}
FUNCTION UDINT_TO_IDENTINGROUP : IDENT_IN_GROUP_REF
VAR_INPUT
	id	:	UDINT;
END_VAR

END_FUNCTION

// POUs/Motion/MC_MovePath

{attribute 'c++_compatible'}
{attribute 'external_name' := 'MC_MovePath_GUID_910966B4_00A6_3665_CD7F_8475FE6F84C3'}
{attribute 'TcIecLibraryType'}
{attribute 'hide_all_locals'}
FUNCTION_BLOCK MC_MovePath
VAR_IN_OUT
	(* B *)
	{attribute 'GUID' := 'EE658783-7533-4695-9194-9C08CBE11A9C'}
	{attribute 'Namespace' := 'Tc3_McCoordinatedMotion'}
	AxesGroup : AXES_GROUP_REF;
	(* B *)
	{attribute 'GUID' := 'C9AD990F-1976-3217-E176-0481FCAF8F1C'}
	{attribute 'Namespace' := 'Tc3_McCoordinatedMotion'}
	PathData : MC_PATH_DATA_REF;
END_VAR
VAR_INPUT
	(* B *)
	Execute : BOOL;
END_VAR
VAR_OUTPUT
	(* B *)
	Done : BOOL;
	(* E *)
	Busy : BOOL;
	(* E *)
	Active : BOOL;
	(* E *)
	CommandAborted : BOOL;
	(* B *)
	Error : BOOL;
END_VAR
VAR
	 {attribute 'hide'}
	_reserved1 : UINT;
END_VAR
VAR_OUTPUT
	(* E *)
	ErrorId : UDINT;
END_VAR
VAR
	 {attribute 'hide'}
	_reserved2 : UINT_0_32;
	InternalFBState : ARRAY [1..16] OF ULINT;
END_VAR

{attribute 'TcTypeSystem'}

(* Internal method *)
{attribute 'hide'}
METHOD FB_init : BOOL
VAR_INPUT
	(*  if TRUE, the retain variables are initialized (warm start / cold start) *)
	bInitRetains : BOOL;
	(*  if TRUE, the instance afterwards gets moved into the copy code (online change) *)
	bInCopyCode : BOOL;
END_VAR
END_METHOD

{attribute 'TcTypeSystem'}

(* Internal method *)
{attribute 'hide'}
METHOD FB_exit : BOOL
VAR_INPUT
	(*  if TRUE, the exit method is called for exiting an instance that is copied afterwards (online change). *)
	bInCopyCode : BOOL;
END_VAR
END_METHOD

END_FUNCTION_BLOCK

// POUs/Motion/MC_BlockerPreparation

{attribute 'c++_compatible'}
{attribute 'external_name' := 'MC_BlockerPreparation_GUID_89150637_2910_36B2_C7FD_D83F8F51DFAD'}
{attribute 'TcIecLibraryType'}
{attribute 'hide_all_locals'}
FUNCTION_BLOCK MC_BlockerPreparation
VAR_IN_OUT
	(* B *)
	{attribute 'GUID' := 'C9AD990F-1976-3217-E176-0481FCAF8F1C'}
	{attribute 'Namespace' := 'Tc3_McCoordinatedMotion'}
	PathData : MC_PATH_DATA_REF;
END_VAR
VAR_INPUT
	(* B *)
	BlockerId : UDINT;
	(* B *)
	{attribute 'Namespace' := 'Tc3_Mc3Definitions'}
	BufferMode : Tc3_Mc3Definitions.MC_BUFFER_MODE;
END_VAR
VAR
	 {attribute 'hide'}
	_reserved1 : UINT;
END_VAR
VAR_INPUT
	(* B *)
	InvokeId : UDINT;
END_VAR
VAR_OUTPUT
	(* B *)
	Error : BOOL;
END_VAR
VAR
	 {attribute 'hide'}
	_reserved2 : ARRAY [1..3] OF USINT;
END_VAR
VAR_OUTPUT
	(* E *)
	ErrorId : UDINT;
END_VAR
VAR
END_VAR

{attribute 'TcTypeSystem'}

(* Internal method *)
{attribute 'hide'}
METHOD FB_init : BOOL
VAR_INPUT
	(*  if TRUE, the retain variables are initialized (warm start / cold start) *)
	bInitRetains : BOOL;
	(*  if TRUE, the instance afterwards gets moved into the copy code (online change) *)
	bInCopyCode : BOOL;
END_VAR
END_METHOD

{attribute 'TcTypeSystem'}

(* Internal method *)
{attribute 'hide'}
METHOD FB_exit : BOOL
VAR_INPUT
	(*  if TRUE, the exit method is called for exiting an instance that is copied afterwards (online change). *)
	bInCopyCode : BOOL;
END_VAR
END_METHOD

END_FUNCTION_BLOCK

// POUs/Motion/MC_DwellTimePreparation

{attribute 'c++_compatible'}
{attribute 'external_name' := 'MC_DwellTimePreparation_GUID_CCC774A8_C834_36C1_F54D_89D0EBBE39FC'}
{attribute 'TcIecLibraryType'}
{attribute 'hide_all_locals'}
FUNCTION_BLOCK MC_DwellTimePreparation
VAR_IN_OUT
	(* B *)
	{attribute 'GUID' := 'C9AD990F-1976-3217-E176-0481FCAF8F1C'}
	{attribute 'Namespace' := 'Tc3_McCoordinatedMotion'}
	PathData : MC_PATH_DATA_REF;
END_VAR
VAR_INPUT
	(* B *)
	DwellTime : TIME;
	(* B *)
	{attribute 'Namespace' := 'Tc3_Mc3Definitions'}
	BufferMode : Tc3_Mc3Definitions.MC_BUFFER_MODE;
END_VAR
VAR
	 {attribute 'hide'}
	_reserved1 : UINT;
END_VAR
VAR_INPUT
	(* B *)
	InvokeId : UDINT;
END_VAR
VAR_OUTPUT
	(* B *)
	Error : BOOL;
END_VAR
VAR
	 {attribute 'hide'}
	_reserved2 : ARRAY [1..3] OF USINT;
END_VAR
VAR_OUTPUT
	(* E *)
	ErrorId : UDINT;
END_VAR
VAR
END_VAR

{attribute 'TcTypeSystem'}

(* Internal method *)
{attribute 'hide'}
METHOD FB_init : BOOL
VAR_INPUT
	(*  if TRUE, the retain variables are initialized (warm start / cold start) *)
	bInitRetains : BOOL;
	(*  if TRUE, the instance afterwards gets moved into the copy code (online change) *)
	bInCopyCode : BOOL;
END_VAR
END_METHOD

{attribute 'TcTypeSystem'}

(* Internal method *)
{attribute 'hide'}
METHOD FB_exit : BOOL
VAR_INPUT
	(*  if TRUE, the exit method is called for exiting an instance that is copied afterwards (online change). *)
	bInCopyCode : BOOL;
END_VAR
END_METHOD

END_FUNCTION_BLOCK

// POUs/Motion/MC_GroupHalt

{attribute 'c++_compatible'}
{attribute 'external_name' := 'MC_GroupHalt_GUID_680BEFB1_DD08_30F3_C8B0_022B23C05D62'}
{attribute 'TcIecLibraryType'}
{attribute 'hide_all_locals'}
FUNCTION_BLOCK MC_GroupHalt
VAR_IN_OUT
	(* B *)
	{attribute 'GUID' := 'EE658783-7533-4695-9194-9C08CBE11A9C'}
	{attribute 'Namespace' := 'Tc3_McCoordinatedMotion'}
	AxesGroup : AXES_GROUP_REF;
END_VAR
VAR_INPUT
	(* B *)
	Execute : BOOL;
END_VAR
VAR
	 {attribute 'hide'}
	_reserved1 : ARRAY [1..7] OF USINT;
END_VAR
VAR_INPUT
	(* E *)
	{attribute 'GUID' := '0100FF8A-3F83-4535-990A-614CFBA4DA63'}
	{attribute 'Namespace' := 'MC'}
	Deceleration : MC.MC_LREAL;
	(* E *)
	{attribute 'GUID' := '0100FF8A-3F83-4535-990A-614CFBA4DA63'}
	{attribute 'Namespace' := 'MC'}
	Jerk : MC.MC_LREAL;
END_VAR
VAR_OUTPUT
	(* E *)
	Done : BOOL;
	(* E *)
	Busy : BOOL;
	(* E *)
	Active : BOOL;
	(* E *)
	CommandAborted : BOOL;
	(* B *)
	Error : BOOL;
END_VAR
VAR
	 {attribute 'hide'}
	_reserved2 : ARRAY [1..3] OF USINT;
END_VAR
VAR_OUTPUT
	(* E *)
	ErrorId : UDINT;
END_VAR
VAR
	 {attribute 'hide'}
	_reserved3 : UDINT;
	InternalFBState : ARRAY [1..16] OF ULINT;
END_VAR

{attribute 'TcTypeSystem'}

(* Internal method *)
{attribute 'hide'}
METHOD FB_init : BOOL
VAR_INPUT
	(*  if TRUE, the retain variables are initialized (warm start / cold start) *)
	bInitRetains : BOOL;
	(*  if TRUE, the instance afterwards gets moved into the copy code (online change) *)
	bInCopyCode : BOOL;
END_VAR
END_METHOD

{attribute 'TcTypeSystem'}

(* Internal method *)
{attribute 'hide'}
METHOD FB_exit : BOOL
VAR_INPUT
	(*  if TRUE, the exit method is called for exiting an instance that is copied afterwards (online change). *)
	bInCopyCode : BOOL;
END_VAR
END_METHOD

END_FUNCTION_BLOCK

// POUs/Motion/MC_GroupStop

{attribute 'c++_compatible'}
{attribute 'external_name' := 'MC_GroupStop_GUID_E2988D5F_9C73_3DEA_CDEA_046D376F5510'}
{attribute 'TcIecLibraryType'}
{attribute 'hide_all_locals'}
FUNCTION_BLOCK MC_GroupStop
VAR_IN_OUT
	(* B *)
	{attribute 'GUID' := 'EE658783-7533-4695-9194-9C08CBE11A9C'}
	{attribute 'Namespace' := 'Tc3_McCoordinatedMotion'}
	AxesGroup : AXES_GROUP_REF;
END_VAR
VAR_INPUT
	(* B *)
	Execute : BOOL;
END_VAR
VAR
	 {attribute 'hide'}
	_reserved1 : ARRAY [1..7] OF USINT;
END_VAR
VAR_INPUT
	(* E *)
	{attribute 'GUID' := '0100FF8A-3F83-4535-990A-614CFBA4DA63'}
	{attribute 'Namespace' := 'MC'}
	Deceleration : MC.MC_LREAL;
	(* E *)
	{attribute 'GUID' := '0100FF8A-3F83-4535-990A-614CFBA4DA63'}
	{attribute 'Namespace' := 'MC'}
	Jerk : MC.MC_LREAL;
END_VAR
VAR_OUTPUT
	(* E *)
	Done : BOOL;
	(* E *)
	Busy : BOOL;
	(* E *)
	Active : BOOL;
	(* E *)
	CommandAborted : BOOL;
	(* B *)
	Error : BOOL;
END_VAR
VAR
	 {attribute 'hide'}
	_reserved2 : ARRAY [1..3] OF USINT;
END_VAR
VAR_OUTPUT
	(* E *)
	ErrorId : UDINT;
END_VAR
VAR
	 {attribute 'hide'}
	_reserved3 : UDINT;
	InternalFBState : ARRAY [1..16] OF ULINT;
END_VAR

{attribute 'TcTypeSystem'}

(* Internal method *)
{attribute 'hide'}
METHOD FB_init : BOOL
VAR_INPUT
	(*  if TRUE, the retain variables are initialized (warm start / cold start) *)
	bInitRetains : BOOL;
	(*  if TRUE, the instance afterwards gets moved into the copy code (online change) *)
	bInCopyCode : BOOL;
END_VAR
END_METHOD

{attribute 'TcTypeSystem'}

(* Internal method *)
{attribute 'hide'}
METHOD FB_exit : BOOL
VAR_INPUT
	(*  if TRUE, the exit method is called for exiting an instance that is copied afterwards (online change). *)
	bInCopyCode : BOOL;
END_VAR
END_METHOD

END_FUNCTION_BLOCK

// POUs/Motion/MC_MoveBlendingPreparation

{attribute 'c++_compatible'}
{attribute 'external_name' := 'MC_MoveBlendingPreparation_GUID_2F60A5E1_7321_335E_F8F1_B920FA04CF11'}
{attribute 'TcIecLibraryType'}
{attribute 'hide_all_locals'}
FUNCTION_BLOCK MC_MoveBlendingPreparation
VAR_IN_OUT
	(* B *)
	{attribute 'GUID' := 'C9AD990F-1976-3217-E176-0481FCAF8F1C'}
	{attribute 'Namespace' := 'Tc3_McCoordinatedMotion'}
	PathData : MC_PATH_DATA_REF;
END_VAR
VAR_INPUT
	(* E *)
	{attribute 'GUID' := '0100FF8A-3F83-4535-990A-614CFBA4DA63'}
	{attribute 'Namespace' := 'MC'}
	Velocity : MC.MC_LREAL;
	(* E *)
	{attribute 'GUID' := '0100FF8A-3F83-4535-990A-614CFBA4DA63'}
	{attribute 'Namespace' := 'MC'}
	Acceleration : MC.MC_LREAL;
	(* E *)
	{attribute 'GUID' := '0100FF8A-3F83-4535-990A-614CFBA4DA63'}
	{attribute 'Namespace' := 'MC'}
	Deceleration : MC.MC_LREAL;
	(* E *)
	{attribute 'GUID' := '0100FF8A-3F83-4535-990A-614CFBA4DA63'}
	{attribute 'Namespace' := 'MC'}
	Jerk : MC.MC_LREAL;
	(* E *)
	{attribute 'Namespace' := 'Tc3_Mc3Definitions'}
	BufferMode : Tc3_Mc3Definitions.MC_BUFFER_MODE;
	(* E *)
	{attribute 'GUID' := 'D5C3E4F6-A7B8-4C9D-AE1F-2A3B4C5D6E7F'}
	{attribute 'Namespace' := 'Tc3_McCoordinatedMotion'}
	TransitionMode : MC_TRANSITION_MODE;
END_VAR
VAR
	 {attribute 'hide'}
	_reserved1 : UINT_0_32;
END_VAR
VAR_INPUT
	(* E *)
	{attribute 'GUID' := '18071995-0000-0000-0000-000000000018'}
	TransitionParameter : GLOBAL.PVOID;
	(* B *)
	TransitionParameterCount : UDINT;
	(* B *)
	InvokeId : UDINT;
	(* E *)
	{attribute 'GUID' := 'B9387A9F-D0A2-9E44-D9DC-1B7D4B662D8E'}
	{attribute 'Namespace' := 'Tc3_Physics'}
	DynamicConstraints : REFERENCE TO Tc3_Physics.IPlcDynamicConstraint;
END_VAR
VAR_OUTPUT
	(* B *)
	Error : BOOL;
END_VAR
VAR
	 {attribute 'hide'}
	_reserved2 : ARRAY [1..3] OF USINT;
END_VAR
VAR_OUTPUT
	(* E *)
	ErrorId : UDINT;
END_VAR
VAR
END_VAR

{attribute 'TcTypeSystem'}

(* Internal method *)
{attribute 'hide'}
METHOD FB_init : BOOL
VAR_INPUT
	(*  if TRUE, the retain variables are initialized (warm start / cold start) *)
	bInitRetains : BOOL;
	(*  if TRUE, the instance afterwards gets moved into the copy code (online change) *)
	bInCopyCode : BOOL;
END_VAR
END_METHOD

{attribute 'TcTypeSystem'}

(* Internal method *)
{attribute 'hide'}
METHOD FB_exit : BOOL
VAR_INPUT
	(*  if TRUE, the exit method is called for exiting an instance that is copied afterwards (online change). *)
	bInCopyCode : BOOL;
END_VAR
END_METHOD

END_FUNCTION_BLOCK

// POUs/Motion/MC_MoveCircularAbsolutePreparation

{attribute 'c++_compatible'}
{attribute 'external_name' := 'MC_MoveCircularAbsolutePreparation_GUID_50CE44DF_9FDB_33F2_DE6B_3EBAF077B487'}
{attribute 'TcIecLibraryType'}
{attribute 'hide_all_locals'}
FUNCTION_BLOCK MC_MoveCircularAbsolutePreparation
VAR_IN_OUT
	(* B *)
	{attribute 'GUID' := 'C9AD990F-1976-3217-E176-0481FCAF8F1C'}
	{attribute 'Namespace' := 'Tc3_McCoordinatedMotion'}
	PathData : MC_PATH_DATA_REF;
END_VAR
VAR_INPUT
	(* B *)
	{attribute 'GUID' := 'B3A1C2D4-E5F6-4A7B-8C9D-0E1F2A3B4C5D'}
	{attribute 'Namespace' := 'Tc3_McCoordinatedMotion'}
	CircMode : MC_CIRC_MODE;
END_VAR
VAR
	 {attribute 'hide'}
	_reserved1 : UINT_16_48;
END_VAR
VAR_INPUT
	(* B *)
	{attribute 'GUID' := '18071995-0000-0000-0000-000000000018'}
	AuxPoint : GLOBAL.PVOID;
	(* B *)
	AuxPointCount : UDINT;
END_VAR
VAR
	 {attribute 'hide'}
	_reserved2 : UINT_0_32;
END_VAR
VAR_INPUT
	(* B *)
	{attribute 'GUID' := '18071995-0000-0000-0000-000000000018'}
	EndPoint : GLOBAL.PVOID;
	(* B *)
	EndPointCount : UDINT;
	(* B *)
	{attribute 'GUID' := 'C4B2D3E5-F6A7-4B8C-9D0E-1F2A3B4C5D6E'}
	{attribute 'Namespace' := 'Tc3_McCoordinatedMotion'}
	PathChoice : MC_CIRC_PATHCHOICE;
END_VAR
VAR
	 {attribute 'hide'}
	_reserved3 : UINT;
END_VAR
VAR_INPUT
	(* E *)
	{attribute 'GUID' := '0100FF8A-3F83-4535-990A-614CFBA4DA63'}
	{attribute 'Namespace' := 'MC'}
	Velocity : MC.MC_LREAL;
	(* E *)
	{attribute 'GUID' := '0100FF8A-3F83-4535-990A-614CFBA4DA63'}
	{attribute 'Namespace' := 'MC'}
	Acceleration : MC.MC_LREAL;
	(* E *)
	{attribute 'GUID' := '0100FF8A-3F83-4535-990A-614CFBA4DA63'}
	{attribute 'Namespace' := 'MC'}
	Deceleration : MC.MC_LREAL;
	(* E *)
	{attribute 'GUID' := '0100FF8A-3F83-4535-990A-614CFBA4DA63'}
	{attribute 'Namespace' := 'MC'}
	Jerk : MC.MC_LREAL;
	(* E *)
	{attribute 'Namespace' := 'Tc3_Mc3Definitions'}
	BufferMode : Tc3_Mc3Definitions.MC_BUFFER_MODE;
	(* E *)
	{attribute 'GUID' := 'D5C3E4F6-A7B8-4C9D-AE1F-2A3B4C5D6E7F'}
	{attribute 'Namespace' := 'Tc3_McCoordinatedMotion'}
	TransitionMode : MC_TRANSITION_MODE;
END_VAR
VAR
	 {attribute 'hide'}
	_reserved4 : UINT_0_32;
END_VAR
VAR_INPUT
	(* E *)
	{attribute 'GUID' := '18071995-0000-0000-0000-000000000018'}
	TransitionParameter : GLOBAL.PVOID;
	(* B *)
	TransitionParameterCount : UDINT;
	(* B *)
	InvokeId : UDINT;
	(* E *)
	{attribute 'GUID' := 'B9387A9F-D0A2-9E44-D9DC-1B7D4B662D8E'}
	{attribute 'Namespace' := 'Tc3_Physics'}
	DynamicConstraints : REFERENCE TO Tc3_Physics.IPlcDynamicConstraint;
END_VAR
VAR_OUTPUT
	(* B *)
	Error : BOOL;
END_VAR
VAR
	 {attribute 'hide'}
	_reserved5 : ARRAY [1..3] OF USINT;
END_VAR
VAR_OUTPUT
	(* E *)
	ErrorId : UDINT;
END_VAR
VAR
END_VAR

{attribute 'TcTypeSystem'}

(* Internal method *)
{attribute 'hide'}
METHOD FB_init : BOOL
VAR_INPUT
	(*  if TRUE, the retain variables are initialized (warm start / cold start) *)
	bInitRetains : BOOL;
	(*  if TRUE, the instance afterwards gets moved into the copy code (online change) *)
	bInCopyCode : BOOL;
END_VAR
END_METHOD

{attribute 'TcTypeSystem'}

(* Internal method *)
{attribute 'hide'}
METHOD FB_exit : BOOL
VAR_INPUT
	(*  if TRUE, the exit method is called for exiting an instance that is copied afterwards (online change). *)
	bInCopyCode : BOOL;
END_VAR
END_METHOD

END_FUNCTION_BLOCK

// POUs/Motion/MC_GroupReadBlockerStatus

{attribute 'c++_compatible'}
{attribute 'external_name' := 'MC_GroupReadBlockerStatus_GUID_0CB62D4F_6DB7_38AF_DFC4_52CB98EACCF2'}
{attribute 'TcIecLibraryType'}
{attribute 'hide_all_locals'}
FUNCTION_BLOCK MC_GroupReadBlockerStatus
VAR_IN_OUT
	(* B *)
	{attribute 'GUID' := 'EE658783-7533-4695-9194-9C08CBE11A9C'}
	{attribute 'Namespace' := 'Tc3_McCoordinatedMotion'}
	AxesGroup : AXES_GROUP_REF;
END_VAR
VAR_INPUT
	(* B *)
	Enable : BOOL;
END_VAR
VAR_OUTPUT
	(* B *)
	Valid : BOOL;
	(* B *)
	Blocked : BOOL;
END_VAR
VAR
	 {attribute 'hide'}
	_reserved1 : USINT;
END_VAR
VAR_OUTPUT
	(* B *)
	BlockerId : UDINT;
END_VAR
VAR
END_VAR

{attribute 'TcTypeSystem'}

(* Internal method *)
{attribute 'hide'}
METHOD FB_init : BOOL
VAR_INPUT
	(*  if TRUE, the retain variables are initialized (warm start / cold start) *)
	bInitRetains : BOOL;
	(*  if TRUE, the instance afterwards gets moved into the copy code (online change) *)
	bInCopyCode : BOOL;
END_VAR
END_METHOD

{attribute 'TcTypeSystem'}

(* Internal method *)
{attribute 'hide'}
METHOD FB_exit : BOOL
VAR_INPUT
	(*  if TRUE, the exit method is called for exiting an instance that is copied afterwards (online change). *)
	bInCopyCode : BOOL;
END_VAR
END_METHOD

END_FUNCTION_BLOCK

// POUs/Motion/MC_MoveDirectPreparation

{attribute 'c++_compatible'}
{attribute 'external_name' := 'MC_MoveDirectPreparation_GUID_64367A38_5BA3_3535_DD1F_8A9F218A99BF'}
{attribute 'TcIecLibraryType'}
{attribute 'hide_all_locals'}
FUNCTION_BLOCK MC_MoveDirectPreparation
VAR_IN_OUT
	(* B *)
	{attribute 'GUID' := 'C9AD990F-1976-3217-E176-0481FCAF8F1C'}
	{attribute 'Namespace' := 'Tc3_McCoordinatedMotion'}
	PathData : MC_PATH_DATA_REF;
END_VAR
VAR_INPUT
	(* B *)
	{attribute 'GUID' := '18071995-0000-0000-0000-000000000018'}
	Position : GLOBAL.PVOID;
	(* B *)
	PositionCount : UDINT;
END_VAR
VAR
	 {attribute 'hide'}
	_reserved1 : UINT_0_32;
END_VAR
VAR_INPUT
	(* E *)
	{attribute 'GUID' := '0100FF8A-3F83-4535-990A-614CFBA4DA63'}
	{attribute 'Namespace' := 'MC'}
	Velocity : MC.MC_LREAL;
	(* E *)
	{attribute 'GUID' := '0100FF8A-3F83-4535-990A-614CFBA4DA63'}
	{attribute 'Namespace' := 'MC'}
	Acceleration : MC.MC_LREAL;
	(* E *)
	{attribute 'GUID' := '0100FF8A-3F83-4535-990A-614CFBA4DA63'}
	{attribute 'Namespace' := 'MC'}
	Deceleration : MC.MC_LREAL;
	(* E *)
	{attribute 'GUID' := '0100FF8A-3F83-4535-990A-614CFBA4DA63'}
	{attribute 'Namespace' := 'MC'}
	Jerk : MC.MC_LREAL;
	(* E *)
	{attribute 'Namespace' := 'Tc3_Mc3Definitions'}
	BufferMode : Tc3_Mc3Definitions.MC_BUFFER_MODE;
	(* E *)
	{attribute 'GUID' := 'D5C3E4F6-A7B8-4C9D-AE1F-2A3B4C5D6E7F'}
	{attribute 'Namespace' := 'Tc3_McCoordinatedMotion'}
	TransitionMode : MC_TRANSITION_MODE;
END_VAR
VAR
	 {attribute 'hide'}
	_reserved2 : UINT_0_32;
END_VAR
VAR_INPUT
	(* E *)
	{attribute 'GUID' := '18071995-0000-0000-0000-000000000018'}
	TransitionParameter : GLOBAL.PVOID;
	(* B *)
	TransitionParameterCount : UDINT;
	(* B *)
	InvokeId : UDINT;
	(* E *)
	{attribute 'GUID' := 'B9387A9F-D0A2-9E44-D9DC-1B7D4B662D8E'}
	{attribute 'Namespace' := 'Tc3_Physics'}
	DynamicConstraints : REFERENCE TO Tc3_Physics.IPlcDynamicConstraint;
END_VAR
VAR_OUTPUT
	(* B *)
	Error : BOOL;
END_VAR
VAR
	 {attribute 'hide'}
	_reserved3 : ARRAY [1..3] OF USINT;
END_VAR
VAR_OUTPUT
	(* E *)
	ErrorId : UDINT;
END_VAR
VAR
END_VAR

{attribute 'TcTypeSystem'}

(* Internal method *)
{attribute 'hide'}
METHOD FB_init : BOOL
VAR_INPUT
	(*  if TRUE, the retain variables are initialized (warm start / cold start) *)
	bInitRetains : BOOL;
	(*  if TRUE, the instance afterwards gets moved into the copy code (online change) *)
	bInCopyCode : BOOL;
END_VAR
END_METHOD

{attribute 'TcTypeSystem'}

(* Internal method *)
{attribute 'hide'}
METHOD FB_exit : BOOL
VAR_INPUT
	(*  if TRUE, the exit method is called for exiting an instance that is copied afterwards (online change). *)
	bInCopyCode : BOOL;
END_VAR
END_METHOD

END_FUNCTION_BLOCK

// POUs/Motion/MC_MoveLinearAbsolutePreparation

{attribute 'c++_compatible'}
{attribute 'external_name' := 'MC_MoveLinearAbsolutePreparation_GUID_5ADEDD70_DC02_3158_E16B_5B09827104B6'}
{attribute 'TcIecLibraryType'}
{attribute 'hide_all_locals'}
FUNCTION_BLOCK MC_MoveLinearAbsolutePreparation
VAR_IN_OUT
	(* B *)
	{attribute 'GUID' := 'C9AD990F-1976-3217-E176-0481FCAF8F1C'}
	{attribute 'Namespace' := 'Tc3_McCoordinatedMotion'}
	PathData : MC_PATH_DATA_REF;
END_VAR
VAR_INPUT
	(* B *)
	{attribute 'GUID' := '18071995-0000-0000-0000-000000000018'}
	Position : GLOBAL.PVOID;
	(* B *)
	PositionCount : UDINT;
END_VAR
VAR
	 {attribute 'hide'}
	_reserved1 : UINT_0_32;
END_VAR
VAR_INPUT
	(* E *)
	{attribute 'GUID' := '0100FF8A-3F83-4535-990A-614CFBA4DA63'}
	{attribute 'Namespace' := 'MC'}
	Velocity : MC.MC_LREAL;
	(* E *)
	{attribute 'GUID' := '0100FF8A-3F83-4535-990A-614CFBA4DA63'}
	{attribute 'Namespace' := 'MC'}
	Acceleration : MC.MC_LREAL;
	(* E *)
	{attribute 'GUID' := '0100FF8A-3F83-4535-990A-614CFBA4DA63'}
	{attribute 'Namespace' := 'MC'}
	Deceleration : MC.MC_LREAL;
	(* E *)
	{attribute 'GUID' := '0100FF8A-3F83-4535-990A-614CFBA4DA63'}
	{attribute 'Namespace' := 'MC'}
	Jerk : MC.MC_LREAL;
	(* E *)
	{attribute 'Namespace' := 'Tc3_Mc3Definitions'}
	BufferMode : Tc3_Mc3Definitions.MC_BUFFER_MODE;
	(* E *)
	{attribute 'GUID' := 'D5C3E4F6-A7B8-4C9D-AE1F-2A3B4C5D6E7F'}
	{attribute 'Namespace' := 'Tc3_McCoordinatedMotion'}
	TransitionMode : MC_TRANSITION_MODE;
END_VAR
VAR
	 {attribute 'hide'}
	_reserved2 : UINT_0_32;
END_VAR
VAR_INPUT
	(* E *)
	{attribute 'GUID' := '18071995-0000-0000-0000-000000000018'}
	TransitionParameter : GLOBAL.PVOID;
	(* B *)
	TransitionParameterCount : UDINT;
	(* B *)
	InvokeId : UDINT;
	(* E *)
	{attribute 'GUID' := 'B9387A9F-D0A2-9E44-D9DC-1B7D4B662D8E'}
	{attribute 'Namespace' := 'Tc3_Physics'}
	DynamicConstraints : REFERENCE TO Tc3_Physics.IPlcDynamicConstraint;
END_VAR
VAR_OUTPUT
	(* B *)
	Error : BOOL;
END_VAR
VAR
	 {attribute 'hide'}
	_reserved3 : ARRAY [1..3] OF USINT;
END_VAR
VAR_OUTPUT
	(* E *)
	ErrorId : UDINT;
END_VAR
VAR
END_VAR

{attribute 'TcTypeSystem'}

(* Internal method *)
{attribute 'hide'}
METHOD FB_init : BOOL
VAR_INPUT
	(*  if TRUE, the retain variables are initialized (warm start / cold start) *)
	bInitRetains : BOOL;
	(*  if TRUE, the instance afterwards gets moved into the copy code (online change) *)
	bInCopyCode : BOOL;
END_VAR
END_METHOD

{attribute 'TcTypeSystem'}

(* Internal method *)
{attribute 'hide'}
METHOD FB_exit : BOOL
VAR_INPUT
	(*  if TRUE, the exit method is called for exiting an instance that is copied afterwards (online change). *)
	bInCopyCode : BOOL;
END_VAR
END_METHOD

END_FUNCTION_BLOCK

// POUs/Motion/MC_ReleaseBlocker

{attribute 'c++_compatible'}
{attribute 'external_name' := 'MC_ReleaseBlocker_GUID_237A98F0_59B2_3E5C_E691_6CAC48697482'}
{attribute 'TcIecLibraryType'}
{attribute 'hide_all_locals'}
FUNCTION_BLOCK MC_ReleaseBlocker
VAR_IN_OUT
	(* B *)
	{attribute 'GUID' := 'EE658783-7533-4695-9194-9C08CBE11A9C'}
	{attribute 'Namespace' := 'Tc3_McCoordinatedMotion'}
	AxesGroup : AXES_GROUP_REF;
END_VAR
VAR_INPUT
	(* B *)
	Execute : BOOL;
END_VAR
VAR
	 {attribute 'hide'}
	_reserved1 : ARRAY [1..3] OF USINT;
END_VAR
VAR_INPUT
	(* E *)
	BlockerId : UDINT;
END_VAR
VAR_OUTPUT
	(* E *)
	Done : BOOL;
	(* E *)
	Busy : BOOL;
	(* B *)
	Error : BOOL;
END_VAR
VAR
	 {attribute 'hide'}
	_reserved2 : USINT;
END_VAR
VAR_OUTPUT
	(* E *)
	ErrorId : UDINT;
END_VAR
VAR
	InternalFBState : ARRAY [1..16] OF ULINT;
END_VAR

{attribute 'TcTypeSystem'}

(* Internal method *)
{attribute 'hide'}
METHOD FB_init : BOOL
VAR_INPUT
	(*  if TRUE, the retain variables are initialized (warm start / cold start) *)
	bInitRetains : BOOL;
	(*  if TRUE, the instance afterwards gets moved into the copy code (online change) *)
	bInCopyCode : BOOL;
END_VAR
END_METHOD

{attribute 'TcTypeSystem'}

(* Internal method *)
{attribute 'hide'}
METHOD FB_exit : BOOL
VAR_INPUT
	(*  if TRUE, the exit method is called for exiting an instance that is copied afterwards (online change). *)
	bInCopyCode : BOOL;
END_VAR
END_METHOD

END_FUNCTION_BLOCK

// POUs/Motion/MC_CalcTrafo

{attribute 'c++_compatible'}
{attribute 'external_name' := 'MC_CalcTrafo_GUID_98D69B44_E078_3CA7_5138_DC89FD59A58D'}
{attribute 'TcIecLibraryType'}
{attribute 'hide_all_locals'}
FUNCTION_BLOCK MC_CalcTrafo
VAR_IN_OUT
	(* B *)
	{attribute 'GUID' := 'EE658783-7533-4695-9194-9C08CBE11A9C'}
	{attribute 'Namespace' := 'Tc3_McCoordinatedMotion'}
	AxesGroup : AXES_GROUP_REF;
	(* E *)
	{attribute 'GUID' := '51DEBB5B-FDCD-4C01-9A10-D37799581013'}
	{attribute 'Namespace' := 'Tc3_McCoordinatedMotion'}
	MetaInfoIn : U_CalcTrafoMetaInfo;
	(* E *)
	{attribute 'GUID' := '51DEBB5B-FDCD-4C01-9A10-D37799581013'}
	{attribute 'Namespace' := 'Tc3_McCoordinatedMotion'}
	MetaInfoOut : U_CalcTrafoMetaInfo;
END_VAR
VAR_INPUT
	(* B *)
	Execute : BOOL;
	(* B *)
	Forward : BOOL;
	(* E *)
	CheckPositionLimits : BOOL := FALSE;
END_VAR
VAR
	 {attribute 'hide'}
	_reserved1 : ARRAY [1..5] OF USINT;
END_VAR
VAR_INPUT
	(* B *)
	AxesPosIn : POINTER TO LREAL;
	(* B *)
	AxesPosInCount : UDINT;
END_VAR
VAR
	 {attribute 'hide'}
	_reserved2 : UINT_0_32;
END_VAR
VAR_INPUT
	(* B *)
	AxesPosOut : POINTER TO LREAL;
	(* B *)
	AxesPosOutCount : UDINT;
END_VAR
VAR_OUTPUT
	(* B *)
	Error : BOOL;
END_VAR
VAR
	 {attribute 'hide'}
	_reserved3 : ARRAY [1..3] OF USINT;
END_VAR
VAR_OUTPUT
	(* E *)
	ErrorId : UDINT;
END_VAR
VAR
	 {attribute 'hide'}
	_reserved4 : UINT_0_32;
END_VAR

{attribute 'TcTypeSystem'}

(* Internal method *)
{attribute 'hide'}
METHOD FB_init : BOOL
VAR_INPUT
	(*  if TRUE, the retain variables are initialized (warm start / cold start) *)
	bInitRetains : BOOL;
	(*  if TRUE, the instance afterwards gets moved into the copy code (online change) *)
	bInCopyCode : BOOL;
END_VAR
END_METHOD

{attribute 'TcTypeSystem'}

(* Internal method *)
{attribute 'hide'}
METHOD FB_exit : BOOL
VAR_INPUT
	(*  if TRUE, the exit method is called for exiting an instance that is copied afterwards (online change). *)
	bInCopyCode : BOOL;
END_VAR
END_METHOD

END_FUNCTION_BLOCK
